(* IEC 61131-3 sources: DigitalTwin/sim-plc/plc, 2 files *)

(* ---- pump_station.st ---- *)
(*
  Pump station lead/lag control: OpenPLC Structured Text program.

  Specification: design/pump-station-design.md, section 4 (logic) and 5 (register map).

  Field I/O (%IX100, %QX100, %IW100) comes from the process simulator, which
  OpenPLC polls as a Modbus "slave device" (Generic TCP, 10.10.0.10:5020).
  The HMI reads the status block %QW0..%QW7 (holding registers 0..7) and
  writes settings to %MW0..%MW10 (holding registers 1024..1034).

  Pressures are UINT scaled x10: 1200 means 120.0 psi.

  Scan order, the same as every PLC: inputs are copied in, this program runs
  top to bottom once, outputs are copied out. Then it starts again.
*)
PROGRAM PumpStation
  VAR
    (* ---- Field inputs from the simulator (design 5.1) ---- *)
    P1_RUNNING    AT %IX100.0 : BOOL;
    P2_RUNNING    AT %IX100.1 : BOOL;
    P1_FAULT      AT %IX100.2 : BOOL;
    P2_FAULT      AT %IX100.3 : BOOL;
    PT101_DISCH   AT %IW100 : UINT;   (* discharge pressure, psi x10 *)
    PT100_SUCT    AT %IW101 : UINT;   (* suction pressure, psi x10 *)
    DEMAND        AT %IW102 : UINT;   (* pipeline demand, % x10 *)
    SIM_HEARTBEAT AT %IW103 : UINT;   (* +1 every simulator step *)

    (* ---- Field outputs to the simulator ---- *)
    P1_RUN_CMD AT %QX100.0 : BOOL;
    P2_RUN_CMD AT %QX100.1 : BOOL;

    (* ---- Status for the HMI: holding registers 0..7 (design 5.2) ---- *)
    HMI_DISCH_PRESS AT %QW0 : UINT;
    HMI_SUCT_PRESS  AT %QW1 : UINT;
    HMI_DEMAND      AT %QW2 : UINT;
    HMI_STATUS      AT %QW3 : UINT;
    HMI_ALARMS      AT %QW4 : UINT;
    HMI_LEAD_PUMP   AT %QW5 : UINT;
    HMI_MODE_ACTIVE AT %QW6 : UINT;
    PLC_HEARTBEAT   AT %QW7 : UINT;

    (* ---- Settings and commands from the HMI: holding registers 1024..1034 (design 5.3) ---- *)
    SP_PRESSURE     AT %MW0 : UINT;   (* lag start pressure, psi x10 *)
    SP_LAG_STOP     AT %MW1 : UINT;   (* lag stop pressure, psi x10 *)
    SP_LOW_ALARM    AT %MW2 : UINT;
    SP_HIGH_ALARM   AT %MW3 : UINT;
    LAG_START_DELAY AT %MW4 : UINT;   (* seconds *)
    LAG_STOP_DELAY  AT %MW5 : UINT;   (* seconds *)
    CMD_MODE        AT %MW6 : UINT;   (* 0 Off, 1 Auto, 2 Manual *)
    CMD_LEAD_SELECT AT %MW7 : UINT;   (* 1 = P1, 2 = P2 *)
    CMD_MANUAL_P1   AT %MW8 : UINT;   (* Manual mode: 1 run, 0 stop *)
    CMD_MANUAL_P2   AT %MW9 : UINT;
    CMD_ALARM_RESET AT %MW10 : UINT;  (* HMI writes 1; the PLC clears it *)
  END_VAR

  VAR
    (* Control state *)
    Mode       : UINT := 0;
    LastMode   : UINT := 0;
    ActiveLead : UINT := 1;        (* lead pump after any failover: 1 or 2 *)
    LagRun     : BOOL := FALSE;    (* Auto logic wants the lag pump running *)
    Handover   : BOOL := FALSE;    (* lead change in progress: keep the old lead on *)
    OldLead    : UINT := 0;
    P1Cmd      : BOOL := FALSE;
    P2Cmd      : BOOL := FALSE;
    LeadRunning : BOOL;
    LagAvail   : BOOL;
    LeadAvail  : BOOL;

    (* Pump failure latches: fault feedback or failed to start. A failed pump
       is locked out (never commanded) until the operator presses Reset and
       the simulator no longer reports a fault. *)
    P1Failed : BOOL := FALSE;
    P2Failed : BOOL := FALSE;
    P1StartTmr : TON;   (* run commanded but no running feedback *)
    P2StartTmr : TON;

    (* Lead/lag timers: the time delays that stop short-cycling *)
    LagStartTmr : TON;
    LagStopTmr  : TON;

    (* Alarms (design 4.3) *)
    LowArmTmr   : TON;   (* start-up bypass for the low-pressure alarm *)
    LowPressTmr : TON;
    HighPressTmr : TON;
    CommLossTmr : TON;
    LastSimHb   : UINT := 0;
    AlmLow   : BOOL := FALSE;
    AlmHigh  : BOOL := FALSE;
    AlmComm  : BOOL := FALSE;
    AlmUnack : BOOL := FALSE;
    AnyAlarm : BOOL;
    PrevAnyAlarm : BOOL := FALSE;
    ResetReq : BOOL;
    CommOk   : BOOL;
    LagRunning : BOOL;
  END_VAR

  (* =====================================================================
     1. First scan: load defaults (design 4.4).
        %MW memory is not kept across a runtime restart, so a zero setpoint
        means "never configured".
     ===================================================================== *)
  IF SP_PRESSURE = 0 THEN
    SP_PRESSURE     := 1200;   (* 120.0 psi *)
    SP_LAG_STOP     := 1450;   (* 145.0 psi *)
    SP_LOW_ALARM    := 1100;   (* 110.0 psi *)
    SP_HIGH_ALARM   := 1600;   (* 160.0 psi *)
    LAG_START_DELAY := 5;
    LAG_STOP_DELAY  := 30;
    CMD_MODE        := 1;      (* Auto *)
    CMD_LEAD_SELECT := 1;      (* P1 *)
    CMD_MANUAL_P1   := 0;
    CMD_MANUAL_P2   := 0;
    CMD_ALARM_RESET := 0;
  END_IF;

  (* =====================================================================
     2. Clamp HMI settings to their allowed ranges (design 5.3).
        The clamped value is written back, so the HMI reads back what the
        PLC is actually using.
     ===================================================================== *)
  SP_PRESSURE := LIMIT(800, SP_PRESSURE, 1500);
  IF SP_LAG_STOP < SP_PRESSURE + 100 THEN
    SP_LAG_STOP := SP_PRESSURE + 100;   (* hysteresis of at least 10 psi *)
  END_IF;
  LAG_START_DELAY := LIMIT(1, LAG_START_DELAY, 60);
  LAG_STOP_DELAY  := LIMIT(5, LAG_STOP_DELAY, 300);
  CMD_MODE        := MIN(CMD_MODE, 2);
  CMD_LEAD_SELECT := LIMIT(1, CMD_LEAD_SELECT, 2);
  CMD_MANUAL_P1   := MIN(CMD_MANUAL_P1, 1);
  CMD_MANUAL_P2   := MIN(CMD_MANUAL_P2, 1);
  Mode := CMD_MODE;

  ResetReq := CMD_ALARM_RESET <> 0;

  (* =====================================================================
     3. Pump health. Fault feedback, or no running feedback 5 s after a run
        command, fails the pump (design 4.2 step 4 and 4.3).
     ===================================================================== *)
  P1StartTmr(IN := P1_RUN_CMD AND NOT P1_RUNNING, PT := T#5s);
  P2StartTmr(IN := P2_RUN_CMD AND NOT P2_RUNNING, PT := T#5s);
  IF P1_FAULT OR P1StartTmr.Q THEN P1Failed := TRUE; END_IF;
  IF P2_FAULT OR P2StartTmr.Q THEN P2Failed := TRUE; END_IF;
  IF ResetReq AND NOT P1_FAULT THEN P1Failed := FALSE; END_IF;
  IF ResetReq AND NOT P2_FAULT THEN P2Failed := FALSE; END_IF;

  (* =====================================================================
     4. Pump control by mode (design 4.1, 4.2)
     ===================================================================== *)
  IF Mode = 1 THEN
    (* ---------------- Auto: lead/lag ---------------- *)

    (* Entering Auto: take the operator's lead choice, and keep whatever
       is already running so the switch causes no bump. *)
    IF LastMode <> 1 THEN
      ActiveLead := CMD_LEAD_SELECT;
      IF ActiveLead = 1 THEN LagRun := P2Cmd; ELSE LagRun := P1Cmd; END_IF;
      Handover := FALSE;
    END_IF;

    (* Failover: the lead pump has failed and the other one is healthy, so
       promote it. The HMI lead selection follows, so the station does not
       swap back on its own once the failed pump is reset. *)
    IF ((ActiveLead = 1) AND P1Failed AND NOT P2Failed) OR
       ((ActiveLead = 2) AND P2Failed AND NOT P1Failed) THEN
      ActiveLead := 3 - ActiveLead;
      CMD_LEAD_SELECT := ActiveLead;
      LagRun := FALSE;
      Handover := FALSE;
    END_IF;

    (* Operator changed the lead pump: applied only while the lag pump is
       stopped (design 4.2 step 5). The old lead keeps running until the new
       one reports running, so pressure does not dip during the swap. *)
    IF (CMD_LEAD_SELECT <> ActiveLead) AND NOT LagRun AND NOT Handover THEN
      IF ((CMD_LEAD_SELECT = 1) AND NOT P1Failed) OR
         ((CMD_LEAD_SELECT = 2) AND NOT P2Failed) THEN
        OldLead := ActiveLead;
        ActiveLead := CMD_LEAD_SELECT;
        Handover := TRUE;
      END_IF;
    END_IF;

    IF ActiveLead = 1 THEN
      LeadAvail := NOT P1Failed;  LagAvail := NOT P2Failed;  LeadRunning := P1_RUNNING;
    ELSE
      LeadAvail := NOT P2Failed;  LagAvail := NOT P1Failed;  LeadRunning := P2_RUNNING;
    END_IF;

    IF Handover AND (LeadRunning OR NOT LeadAvail) THEN
      Handover := FALSE;
    END_IF;

    (* Lag start: pressure below setpoint for the start delay (step 2) *)
    LagStartTmr(IN := (PT101_DISCH < SP_PRESSURE) AND NOT LagRun AND LagAvail AND NOT Handover,
                PT := T#1s * UINT_TO_DINT(LAG_START_DELAY));
    IF LagStartTmr.Q THEN
      LagRun := TRUE;
    END_IF;

    (* Lag stop: pressure above the lag stop pressure for the stop delay (step 3).
       The gap between 120 and 145 psi is the hysteresis that stops cycling. *)
    LagStopTmr(IN := LagRun AND (PT101_DISCH > SP_LAG_STOP),
               PT := T#1s * UINT_TO_DINT(LAG_STOP_DELAY));
    IF LagStopTmr.Q OR NOT LagAvail THEN
      LagRun := FALSE;
    END_IF;

    (* Lead always runs (step 1); lag runs when called for *)
    IF ActiveLead = 1 THEN
      P1Cmd := TRUE;
      P2Cmd := LagRun OR (Handover AND OldLead = 2);
    ELSE
      P2Cmd := TRUE;
      P1Cmd := LagRun OR (Handover AND OldLead = 1);
    END_IF;

  ELSIF Mode = 2 THEN
    (* ---------------- Manual: operator runs each pump ---------------- *)
    P1Cmd := CMD_MANUAL_P1 = 1;
    P2Cmd := CMD_MANUAL_P2 = 1;
    LagRun := FALSE;
    Handover := FALSE;

  ELSE
    (* ---------------- Off ---------------- *)
    P1Cmd := FALSE;
    P2Cmd := FALSE;
    LagRun := FALSE;
    Handover := FALSE;
  END_IF;

  (* Interlock in every mode: a failed pump is never commanded *)
  IF P1Failed THEN P1Cmd := FALSE; END_IF;
  IF P2Failed THEN P2Cmd := FALSE; END_IF;
  P1_RUN_CMD := P1Cmd;
  P2_RUN_CMD := P2Cmd;

  (* Outside Manual, the manual commands track the pumps, so switching to
     Manual leaves them as they are (bumpless transfer). *)
  IF Mode <> 2 THEN
    CMD_MANUAL_P1 := BOOL_TO_UINT(P1Cmd);
    CMD_MANUAL_P2 := BOOL_TO_UINT(P2Cmd);
  END_IF;
  LastMode := Mode;

  (* =====================================================================
     5. Alarms (design 4.3). Each one latches until the operator presses
        Reset AND its condition has cleared.
     ===================================================================== *)

  (* Low pressure is armed once the station has been out of Off for 15 s,
     so a normal start-up (pressure rising from 20 psi) does not alarm. *)
  LowArmTmr(IN := Mode <> 0, PT := T#15s);
  LowPressTmr(IN := LowArmTmr.Q AND (PT101_DISCH < SP_LOW_ALARM), PT := T#5s);
  HighPressTmr(IN := PT101_DISCH > SP_HIGH_ALARM, PT := T#5s);

  (* Simulator comm loss: heartbeat has not changed for 3 s *)
  CommLossTmr(IN := SIM_HEARTBEAT = LastSimHb, PT := T#3s);
  LastSimHb := SIM_HEARTBEAT;
  CommOk := NOT CommLossTmr.Q;

  IF LowPressTmr.Q  THEN AlmLow  := TRUE; END_IF;
  IF HighPressTmr.Q THEN AlmHigh := TRUE; END_IF;
  IF CommLossTmr.Q  THEN AlmComm := TRUE; END_IF;

  IF ResetReq THEN
    IF NOT LowPressTmr.Q  THEN AlmLow  := FALSE; END_IF;
    IF NOT HighPressTmr.Q THEN AlmHigh := FALSE; END_IF;
    IF NOT CommLossTmr.Q  THEN AlmComm := FALSE; END_IF;
    AlmUnack := FALSE;          (* Reset also acknowledges *)
    CMD_ALARM_RESET := 0;       (* handled *)
  END_IF;

  (* A newly raised alarm is unacknowledged until the next Reset *)
  AnyAlarm := AlmLow OR AlmHigh OR P1Failed OR P2Failed OR AlmComm;
  IF AnyAlarm AND NOT PrevAnyAlarm THEN AlmUnack := TRUE; END_IF;
  PrevAnyAlarm := AnyAlarm;

  (* =====================================================================
     6. Status block for the HMI (design 5.2)
     ===================================================================== *)
  IF ActiveLead = 1 THEN LagRunning := P2_RUNNING; ELSE LagRunning := P1_RUNNING; END_IF;

  HMI_DISCH_PRESS := PT101_DISCH;
  HMI_SUCT_PRESS  := PT100_SUCT;
  HMI_DEMAND      := DEMAND;
  HMI_STATUS := BOOL_TO_UINT(P1_RUN_CMD)
              + BOOL_TO_UINT(P1_RUNNING) * 2
              + BOOL_TO_UINT(P2_RUN_CMD) * 4
              + BOOL_TO_UINT(P2_RUNNING) * 8
              + BOOL_TO_UINT(LagRunning) * 16
              + BOOL_TO_UINT(CommOk)     * 32;
  HMI_ALARMS := BOOL_TO_UINT(AlmLow)
              + BOOL_TO_UINT(AlmHigh)  * 2
              + BOOL_TO_UINT(P1Failed) * 4
              + BOOL_TO_UINT(P2Failed) * 8
              + BOOL_TO_UINT(AlmComm)  * 16
              + BOOL_TO_UINT(AlmUnack) * 32768;
  HMI_LEAD_PUMP   := ActiveLead;
  HMI_MODE_ACTIVE := Mode;

  IF PLC_HEARTBEAT = 65535 THEN
    PLC_HEARTBEAT := 0;
  ELSE
    PLC_HEARTBEAT := PLC_HEARTBEAT + 1;
  END_IF;
END_PROGRAM

CONFIGURATION Config0
  RESOURCE Res0 ON PLC
    TASK MainTask(INTERVAL := T#100ms, PRIORITY := 0);
    PROGRAM Inst0 WITH MainTask : PumpStation;
  END_RESOURCE
END_CONFIGURATION

(* ---- pump_station_ld.st ---- *)
(*
  Generated from the ladder program in pump_station_ld/plc.xml by OpenPLC Editor's
  code generator. Do not edit this file: change the ladder in OpenPLC Editor instead.

  Upload this file to OpenPLC Runtime (Programs -> Upload program), or run
      python3 deploy_to_openplc.py --program pump_station_ld.st
  It behaves exactly like pump_station.st and uses the same register map.
*)
PROGRAM PumpStation
  VAR
    LoadDefaults : BOOL;
    MinLagStop : UINT;
    ModeAuto : BOOL;
    ModeManual : BOOL;
    SelP2 : BOOL;
    ManP1 : BOOL;
    ManP2 : BOOL;
    ResetReq : BOOL;
    PressBelowSP : BOOL;
    PressAboveLagStop : BOOL;
    PressBelowLowAlm : BOOL;
    PressAboveHighAlm : BOOL;
    P1StartTmr : TON;
    P2StartTmr : TON;
    P1StartFail : BOOL;
    P2StartFail : BOOL;
    P1Failed : BOOL;
    P2Failed : BOOL;
    EnterAuto : BOOL;
    LeadIsP2 : BOOL;
    LagPumpCmd : BOOL;
    FailToP2 : BOOL;
    FailToP1 : BOOL;
    LeadChange : BOOL;
    LagRun : BOOL;
    Handover : BOOL;
    LeadAvail : BOOL;
    LagAvail : BOOL;
    LeadRunning : BOOL;
    LagStartPT : TIME;
    LagStopPT : TIME;
    LagStartTmr : TON;
    LagStopTmr : TON;
    LagStartDone : BOOL;
    LagStopDone : BOOL;
    LowArmTmr : TON;
    LowPressTmr : TON;
    HighPressTmr : TON;
    CommLossTmr : TON;
    LowArmed : BOOL;
    LowPressOn : BOOL;
    HighPressOn : BOOL;
    SimHbFrozen : BOOL;
    LastSimHb : UINT;
    CommLost : BOOL;
    CommOk : BOOL;
    AlmLow : BOOL;
    AlmHigh : BOOL;
    AlmComm : BOOL;
    AlmUnack : BOOL;
    AnyAlarm : BOOL;
    LagRunning : BOOL;
    StatusWord : UINT;
    AlarmWord : UINT;
    HbWrap : BOOL;
  END_VAR
  VAR
    P1_RUNNING AT %IX100.0 : BOOL;
    P2_RUNNING AT %IX100.1 : BOOL;
    P1_FAULT AT %IX100.2 : BOOL;
    P2_FAULT AT %IX100.3 : BOOL;
    PT101_DISCH AT %IW100 : UINT;
    PT100_SUCT AT %IW101 : UINT;
    DEMAND AT %IW102 : UINT;
    SIM_HEARTBEAT AT %IW103 : UINT;
    P1_RUN_CMD AT %QX100.0 : BOOL;
    P2_RUN_CMD AT %QX100.1 : BOOL;
    HMI_DISCH_PRESS AT %QW0 : UINT;
    HMI_SUCT_PRESS AT %QW1 : UINT;
    HMI_DEMAND AT %QW2 : UINT;
    HMI_STATUS AT %QW3 : UINT;
    HMI_ALARMS AT %QW4 : UINT;
    HMI_LEAD_PUMP AT %QW5 : UINT;
    HMI_MODE_ACTIVE AT %QW6 : UINT;
    PLC_HEARTBEAT AT %QW7 : UINT;
    SP_PRESSURE AT %MW0 : UINT;
    SP_LAG_STOP AT %MW1 : UINT;
    SP_LOW_ALARM AT %MW2 : UINT;
    SP_HIGH_ALARM AT %MW3 : UINT;
    LAG_START_DELAY AT %MW4 : UINT;
    LAG_STOP_DELAY AT %MW5 : UINT;
    CMD_MODE AT %MW6 : UINT;
    CMD_LEAD_SELECT AT %MW7 : UINT;
    CMD_MANUAL_P1 AT %MW8 : UINT;
    CMD_MANUAL_P2 AT %MW9 : UINT;
    CMD_ALARM_RESET AT %MW10 : UINT;
  END_VAR
  VAR
    _TMP_EQ5_OUT : BOOL;
    _TMP_MOVE11_ENO : BOOL;
    _TMP_MOVE11_OUT : UINT;
    _TMP_MOVE14_ENO : BOOL;
    _TMP_MOVE14_OUT : UINT;
    _TMP_MOVE17_ENO : BOOL;
    _TMP_MOVE17_OUT : UINT;
    _TMP_MOVE20_ENO : BOOL;
    _TMP_MOVE20_OUT : UINT;
    _TMP_MOVE23_ENO : BOOL;
    _TMP_MOVE23_OUT : UINT;
    _TMP_MOVE26_ENO : BOOL;
    _TMP_MOVE26_OUT : UINT;
    _TMP_MOVE29_ENO : BOOL;
    _TMP_MOVE29_OUT : UINT;
    _TMP_MOVE32_ENO : BOOL;
    _TMP_MOVE32_OUT : UINT;
    _TMP_MOVE35_ENO : BOOL;
    _TMP_MOVE35_OUT : UINT;
    _TMP_MOVE38_ENO : BOOL;
    _TMP_MOVE38_OUT : UINT;
    _TMP_MOVE41_ENO : BOOL;
    _TMP_MOVE41_OUT : UINT;
    _TMP_LIMIT48_ENO : BOOL;
    _TMP_LIMIT48_OUT : UINT;
    _TMP_ADD53_ENO : BOOL;
    _TMP_ADD53_OUT : UINT;
    _TMP_MAX58_ENO : BOOL;
    _TMP_MAX58_OUT : UINT;
    _TMP_LIMIT64_ENO : BOOL;
    _TMP_LIMIT64_OUT : UINT;
    _TMP_LIMIT70_ENO : BOOL;
    _TMP_LIMIT70_OUT : UINT;
    _TMP_MIN76_ENO : BOOL;
    _TMP_MIN76_OUT : UINT;
    _TMP_LIMIT82_ENO : BOOL;
    _TMP_LIMIT82_OUT : UINT;
    _TMP_MIN87_ENO : BOOL;
    _TMP_MIN87_OUT : UINT;
    _TMP_MIN92_ENO : BOOL;
    _TMP_MIN92_OUT : UINT;
    _TMP_EQ98_OUT : BOOL;
    _TMP_EQ102_OUT : BOOL;
    _TMP_EQ107_OUT : BOOL;
    _TMP_EQ111_OUT : BOOL;
    _TMP_EQ115_OUT : BOOL;
    _TMP_NE119_OUT : BOOL;
    _TMP_LT124_OUT : BOOL;
    _TMP_GT128_OUT : BOOL;
    _TMP_LT132_OUT : BOOL;
    _TMP_GT136_OUT : BOOL;
    R_TRIG1 : R_TRIG;
    _TMP_MOVE220_ENO : BOOL;
    _TMP_MOVE220_OUT : UINT;
    _TMP_MOVE227_ENO : BOOL;
    _TMP_MOVE227_OUT : UINT;
    _TMP_UINT_TO_TIME286_ENO : BOOL;
    _TMP_UINT_TO_TIME286_OUT : TIME;
    _TMP_UINT_TO_TIME290_ENO : BOOL;
    _TMP_UINT_TO_TIME290_OUT : TIME;
    _TMP_BOOL_TO_UINT352_ENO : BOOL;
    _TMP_BOOL_TO_UINT352_OUT : UINT;
    _TMP_BOOL_TO_UINT355_ENO : BOOL;
    _TMP_BOOL_TO_UINT355_OUT : UINT;
    _TMP_EQ382_OUT : BOOL;
    _TMP_MOVE390_ENO : BOOL;
    _TMP_MOVE390_OUT : UINT;
    _TMP_MOVE417_ENO : BOOL;
    _TMP_MOVE417_OUT : UINT;
    R_TRIG2 : R_TRIG;
    _TMP_MOVE445_ENO : BOOL;
    _TMP_MOVE445_OUT : UINT;
    _TMP_MOVE449_ENO : BOOL;
    _TMP_MOVE449_OUT : UINT;
    _TMP_MOVE453_ENO : BOOL;
    _TMP_MOVE453_OUT : UINT;
    _TMP_SEL459_ENO : BOOL;
    _TMP_SEL459_OUT : UINT;
    _TMP_MOVE463_ENO : BOOL;
    _TMP_MOVE463_OUT : UINT;
    _TMP_MOVE468_ENO : BOOL;
    _TMP_MOVE468_OUT : UINT;
    _TMP_ADD475_ENO : BOOL;
    _TMP_ADD475_OUT : UINT;
    _TMP_ADD481_ENO : BOOL;
    _TMP_ADD481_OUT : UINT;
    _TMP_ADD487_ENO : BOOL;
    _TMP_ADD487_OUT : UINT;
    _TMP_ADD493_ENO : BOOL;
    _TMP_ADD493_OUT : UINT;
    _TMP_ADD499_ENO : BOOL;
    _TMP_ADD499_OUT : UINT;
    _TMP_ADD505_ENO : BOOL;
    _TMP_ADD505_OUT : UINT;
    _TMP_MOVE508_ENO : BOOL;
    _TMP_MOVE508_OUT : UINT;
    _TMP_MOVE513_ENO : BOOL;
    _TMP_MOVE513_OUT : UINT;
    _TMP_ADD520_ENO : BOOL;
    _TMP_ADD520_OUT : UINT;
    _TMP_ADD526_ENO : BOOL;
    _TMP_ADD526_OUT : UINT;
    _TMP_ADD532_ENO : BOOL;
    _TMP_ADD532_OUT : UINT;
    _TMP_ADD538_ENO : BOOL;
    _TMP_ADD538_OUT : UINT;
    _TMP_ADD544_ENO : BOOL;
    _TMP_ADD544_OUT : UINT;
    _TMP_ADD550_ENO : BOOL;
    _TMP_ADD550_OUT : UINT;
    _TMP_MOVE553_ENO : BOOL;
    _TMP_MOVE553_OUT : UINT;
    _TMP_EQ559_OUT : BOOL;
    _TMP_ADD565_ENO : BOOL;
    _TMP_ADD565_OUT : UINT;
    _TMP_MOVE570_ENO : BOOL;
    _TMP_MOVE570_OUT : UINT;
  END_VAR

  _TMP_EQ5_OUT := EQ(SP_PRESSURE, 0);
  LoadDefaults := _TMP_EQ5_OUT;
  _TMP_MOVE11_OUT := MOVE(EN := LoadDefaults, IN := 1200, ENO => _TMP_MOVE11_ENO);
  IF _TMP_MOVE11_ENO THEN
      SP_PRESSURE := _TMP_MOVE11_OUT;
  END_IF;
  _TMP_MOVE14_OUT := MOVE(EN := LoadDefaults, IN := 1450, ENO => _TMP_MOVE14_ENO);
  IF _TMP_MOVE14_ENO THEN
      SP_LAG_STOP := _TMP_MOVE14_OUT;
  END_IF;
  _TMP_MOVE17_OUT := MOVE(EN := LoadDefaults, IN := 1100, ENO => _TMP_MOVE17_ENO);
  IF _TMP_MOVE17_ENO THEN
      SP_LOW_ALARM := _TMP_MOVE17_OUT;
  END_IF;
  _TMP_MOVE20_OUT := MOVE(EN := LoadDefaults, IN := 1600, ENO => _TMP_MOVE20_ENO);
  IF _TMP_MOVE20_ENO THEN
      SP_HIGH_ALARM := _TMP_MOVE20_OUT;
  END_IF;
  _TMP_MOVE23_OUT := MOVE(EN := LoadDefaults, IN := 5, ENO => _TMP_MOVE23_ENO);
  IF _TMP_MOVE23_ENO THEN
      LAG_START_DELAY := _TMP_MOVE23_OUT;
  END_IF;
  _TMP_MOVE26_OUT := MOVE(EN := LoadDefaults, IN := 30, ENO => _TMP_MOVE26_ENO);
  IF _TMP_MOVE26_ENO THEN
      LAG_STOP_DELAY := _TMP_MOVE26_OUT;
  END_IF;
  _TMP_MOVE29_OUT := MOVE(EN := LoadDefaults, IN := 1, ENO => _TMP_MOVE29_ENO);
  IF _TMP_MOVE29_ENO THEN
      CMD_MODE := _TMP_MOVE29_OUT;
  END_IF;
  _TMP_MOVE32_OUT := MOVE(EN := LoadDefaults, IN := 1, ENO => _TMP_MOVE32_ENO);
  IF _TMP_MOVE32_ENO THEN
      CMD_LEAD_SELECT := _TMP_MOVE32_OUT;
  END_IF;
  _TMP_MOVE35_OUT := MOVE(EN := LoadDefaults, IN := 0, ENO => _TMP_MOVE35_ENO);
  IF _TMP_MOVE35_ENO THEN
      CMD_MANUAL_P1 := _TMP_MOVE35_OUT;
  END_IF;
  _TMP_MOVE38_OUT := MOVE(EN := LoadDefaults, IN := 0, ENO => _TMP_MOVE38_ENO);
  IF _TMP_MOVE38_ENO THEN
      CMD_MANUAL_P2 := _TMP_MOVE38_OUT;
  END_IF;
  _TMP_MOVE41_OUT := MOVE(EN := LoadDefaults, IN := 0, ENO => _TMP_MOVE41_ENO);
  IF _TMP_MOVE41_ENO THEN
      CMD_ALARM_RESET := _TMP_MOVE41_OUT;
  END_IF;
  _TMP_LIMIT48_OUT := LIMIT(EN := TRUE, MN := 800, IN := SP_PRESSURE, MX := 1500, ENO => _TMP_LIMIT48_ENO);
  IF _TMP_LIMIT48_ENO THEN
      SP_PRESSURE := _TMP_LIMIT48_OUT;
  END_IF;
  _TMP_ADD53_OUT := ADD(EN := TRUE, IN1 := SP_PRESSURE, IN2 := 100, ENO => _TMP_ADD53_ENO);
  IF _TMP_ADD53_ENO THEN
      MinLagStop := _TMP_ADD53_OUT;
  END_IF;
  _TMP_MAX58_OUT := MAX(EN := TRUE, IN1 := SP_LAG_STOP, IN2 := MinLagStop, ENO => _TMP_MAX58_ENO);
  IF _TMP_MAX58_ENO THEN
      SP_LAG_STOP := _TMP_MAX58_OUT;
  END_IF;
  _TMP_LIMIT64_OUT := LIMIT(EN := TRUE, MN := 1, IN := LAG_START_DELAY, MX := 60, ENO => _TMP_LIMIT64_ENO);
  IF _TMP_LIMIT64_ENO THEN
      LAG_START_DELAY := _TMP_LIMIT64_OUT;
  END_IF;
  _TMP_LIMIT70_OUT := LIMIT(EN := TRUE, MN := 5, IN := LAG_STOP_DELAY, MX := 300, ENO => _TMP_LIMIT70_ENO);
  IF _TMP_LIMIT70_ENO THEN
      LAG_STOP_DELAY := _TMP_LIMIT70_OUT;
  END_IF;
  _TMP_MIN76_OUT := MIN(EN := TRUE, IN1 := CMD_MODE, IN2 := 2, ENO => _TMP_MIN76_ENO);
  IF _TMP_MIN76_ENO THEN
      CMD_MODE := _TMP_MIN76_OUT;
  END_IF;
  _TMP_LIMIT82_OUT := LIMIT(EN := TRUE, MN := 1, IN := CMD_LEAD_SELECT, MX := 2, ENO => _TMP_LIMIT82_ENO);
  IF _TMP_LIMIT82_ENO THEN
      CMD_LEAD_SELECT := _TMP_LIMIT82_OUT;
  END_IF;
  _TMP_MIN87_OUT := MIN(EN := TRUE, IN1 := CMD_MANUAL_P1, IN2 := 1, ENO => _TMP_MIN87_ENO);
  IF _TMP_MIN87_ENO THEN
      CMD_MANUAL_P1 := _TMP_MIN87_OUT;
  END_IF;
  _TMP_MIN92_OUT := MIN(EN := TRUE, IN1 := CMD_MANUAL_P2, IN2 := 1, ENO => _TMP_MIN92_ENO);
  IF _TMP_MIN92_ENO THEN
      CMD_MANUAL_P2 := _TMP_MIN92_OUT;
  END_IF;
  _TMP_EQ98_OUT := EQ(CMD_MODE, 1);
  ModeAuto := _TMP_EQ98_OUT;
  _TMP_EQ102_OUT := EQ(CMD_MODE, 2);
  ModeManual := _TMP_EQ102_OUT;
  _TMP_EQ107_OUT := EQ(CMD_LEAD_SELECT, 2);
  SelP2 := _TMP_EQ107_OUT;
  _TMP_EQ111_OUT := EQ(CMD_MANUAL_P1, 1);
  ManP1 := _TMP_EQ111_OUT;
  _TMP_EQ115_OUT := EQ(CMD_MANUAL_P2, 1);
  ManP2 := _TMP_EQ115_OUT;
  _TMP_NE119_OUT := NE(CMD_ALARM_RESET, 0);
  ResetReq := _TMP_NE119_OUT;
  _TMP_LT124_OUT := LT(PT101_DISCH, SP_PRESSURE);
  PressBelowSP := _TMP_LT124_OUT;
  _TMP_GT128_OUT := GT(PT101_DISCH, SP_LAG_STOP);
  PressAboveLagStop := _TMP_GT128_OUT;
  _TMP_LT132_OUT := LT(PT101_DISCH, SP_LOW_ALARM);
  PressBelowLowAlm := _TMP_LT132_OUT;
  _TMP_GT136_OUT := GT(PT101_DISCH, SP_HIGH_ALARM);
  PressAboveHighAlm := _TMP_GT136_OUT;
  P1StartTmr(IN := NOT(P1_RUNNING) AND P1_RUN_CMD, PT := T#5s);
  P1StartFail := P1StartTmr.Q;
  P2StartTmr(IN := NOT(P2_RUNNING) AND P2_RUN_CMD, PT := T#5s);
  P2StartFail := P2StartTmr.Q;
  IF P1StartFail OR P1_FAULT THEN
    P1Failed := TRUE; (*set*)
  END_IF;
  IF P2StartFail OR P2_FAULT THEN
    P2Failed := TRUE; (*set*)
  END_IF;
  IF NOT(P1_FAULT) AND ResetReq THEN
    P1Failed := FALSE; (*reset*)
  END_IF;
  IF NOT(P2_FAULT) AND ResetReq THEN
    P2Failed := FALSE; (*reset*)
  END_IF;
  R_TRIG1(CLK := ModeAuto);
  EnterAuto := R_TRIG1.Q;
  IF SelP2 AND EnterAuto THEN
    LeadIsP2 := TRUE; (*set*)
  END_IF;
  IF NOT(SelP2) AND EnterAuto THEN
    LeadIsP2 := FALSE; (*reset*)
  END_IF;
  LagPumpCmd := P1_RUN_CMD AND LeadIsP2 OR P2_RUN_CMD AND NOT(LeadIsP2);
  IF LagPumpCmd AND EnterAuto THEN
    LagRun := TRUE; (*set*)
  END_IF;
  IF NOT(LagPumpCmd) AND EnterAuto THEN
    LagRun := FALSE; (*reset*)
  END_IF;
  IF EnterAuto THEN
    Handover := FALSE; (*reset*)
  END_IF;
  FailToP2 := NOT(P2Failed) AND P1Failed AND NOT(LeadIsP2) AND ModeAuto;
  FailToP1 := NOT(P1Failed) AND P2Failed AND LeadIsP2 AND ModeAuto;
  IF FailToP2 THEN
    LeadIsP2 := TRUE; (*set*)
  END_IF;
  IF FailToP2 THEN
    SelP2 := TRUE; (*set*)
  END_IF;
  _TMP_MOVE220_OUT := MOVE(EN := FailToP2, IN := 2, ENO => _TMP_MOVE220_ENO);
  IF _TMP_MOVE220_ENO THEN
      CMD_LEAD_SELECT := _TMP_MOVE220_OUT;
  END_IF;
  IF FailToP1 THEN
    LeadIsP2 := FALSE; (*reset*)
  END_IF;
  IF FailToP1 THEN
    SelP2 := FALSE; (*reset*)
  END_IF;
  _TMP_MOVE227_OUT := MOVE(EN := FailToP1, IN := 1, ENO => _TMP_MOVE227_ENO);
  IF _TMP_MOVE227_ENO THEN
      CMD_LEAD_SELECT := _TMP_MOVE227_OUT;
  END_IF;
  IF FailToP1 OR FailToP2 THEN
    LagRun := FALSE; (*reset*)
  END_IF;
  IF FailToP1 OR FailToP2 THEN
    Handover := FALSE; (*reset*)
  END_IF;
  LeadChange := (NOT(P2Failed) AND NOT(LeadIsP2) AND SelP2 OR NOT(P1Failed) AND LeadIsP2 AND NOT(SelP2)) AND NOT(Handover) AND NOT(LagRun) AND ModeAuto;
  IF SelP2 AND LeadChange THEN
    LeadIsP2 := TRUE; (*set*)
  END_IF;
  IF NOT(SelP2) AND LeadChange THEN
    LeadIsP2 := FALSE; (*reset*)
  END_IF;
  IF LeadChange THEN
    Handover := TRUE; (*set*)
  END_IF;
  LeadAvail := NOT(P1Failed) AND NOT(LeadIsP2) OR NOT(P2Failed) AND LeadIsP2;
  LagAvail := NOT(P2Failed) AND NOT(LeadIsP2) OR NOT(P1Failed) AND LeadIsP2;
  LeadRunning := P1_RUNNING AND NOT(LeadIsP2) OR P2_RUNNING AND LeadIsP2;
  IF (LeadRunning OR NOT(LeadAvail)) AND Handover AND ModeAuto THEN
    Handover := FALSE; (*reset*)
  END_IF;
  _TMP_UINT_TO_TIME286_OUT := UINT_TO_TIME(EN := TRUE, IN := LAG_START_DELAY, ENO => _TMP_UINT_TO_TIME286_ENO);
  IF _TMP_UINT_TO_TIME286_ENO THEN
      LagStartPT := _TMP_UINT_TO_TIME286_OUT;
  END_IF;
  _TMP_UINT_TO_TIME290_OUT := UINT_TO_TIME(EN := TRUE, IN := LAG_STOP_DELAY, ENO => _TMP_UINT_TO_TIME290_ENO);
  IF _TMP_UINT_TO_TIME290_ENO THEN
      LagStopPT := _TMP_UINT_TO_TIME290_OUT;
  END_IF;
  LagStartTmr(EN := ModeAuto, IN := NOT(Handover) AND LagAvail AND NOT(LagRun) AND PressBelowSP, PT := LagStartPT);
  LagStartDone := LagStartTmr.Q;
  IF LagStartDone AND ModeAuto THEN
    LagRun := TRUE; (*set*)
  END_IF;
  LagStopTmr(EN := ModeAuto, IN := PressAboveLagStop AND LagRun, PT := LagStopPT);
  LagStopDone := LagStopTmr.Q;
  IF (LagStopDone OR NOT(LagAvail)) AND ModeAuto THEN
    LagRun := FALSE; (*reset*)
  END_IF;
  IF NOT(ModeAuto) THEN
    LagRun := FALSE; (*reset*)
  END_IF;
  IF NOT(ModeAuto) THEN
    Handover := FALSE; (*reset*)
  END_IF;
  P1_RUN_CMD := ((Handover OR LagRun OR NOT(LeadIsP2)) AND ModeAuto OR ManP1 AND ModeManual) AND NOT(P1Failed);
  P2_RUN_CMD := ((Handover OR LagRun OR LeadIsP2) AND ModeAuto OR ManP2 AND ModeManual) AND NOT(P2Failed);
  _TMP_BOOL_TO_UINT352_OUT := BOOL_TO_UINT(EN := NOT(ModeManual), IN := P1_RUN_CMD, ENO => _TMP_BOOL_TO_UINT352_ENO);
  IF _TMP_BOOL_TO_UINT352_ENO THEN
      CMD_MANUAL_P1 := _TMP_BOOL_TO_UINT352_OUT;
  END_IF;
  _TMP_BOOL_TO_UINT355_OUT := BOOL_TO_UINT(EN := NOT(ModeManual), IN := P2_RUN_CMD, ENO => _TMP_BOOL_TO_UINT355_ENO);
  IF _TMP_BOOL_TO_UINT355_ENO THEN
      CMD_MANUAL_P2 := _TMP_BOOL_TO_UINT355_OUT;
  END_IF;
  LowArmTmr(IN := ModeAuto OR ModeManual, PT := T#15s);
  LowArmed := LowArmTmr.Q;
  LowPressTmr(IN := PressBelowLowAlm AND LowArmed, PT := T#5s);
  LowPressOn := LowPressTmr.Q;
  HighPressTmr(IN := PressAboveHighAlm, PT := T#5s);
  HighPressOn := HighPressTmr.Q;
  _TMP_EQ382_OUT := EQ(SIM_HEARTBEAT, LastSimHb);
  SimHbFrozen := _TMP_EQ382_OUT;
  CommLossTmr(IN := SimHbFrozen, PT := T#3s);
  CommLost := CommLossTmr.Q;
  _TMP_MOVE390_OUT := MOVE(EN := TRUE, IN := SIM_HEARTBEAT, ENO => _TMP_MOVE390_ENO);
  IF _TMP_MOVE390_ENO THEN
      LastSimHb := _TMP_MOVE390_OUT;
  END_IF;
  CommOk := NOT(CommLost);
  IF LowPressOn THEN
    AlmLow := TRUE; (*set*)
  END_IF;
  IF HighPressOn THEN
    AlmHigh := TRUE; (*set*)
  END_IF;
  IF CommLost THEN
    AlmComm := TRUE; (*set*)
  END_IF;
  IF NOT(LowPressOn) AND ResetReq THEN
    AlmLow := FALSE; (*reset*)
  END_IF;
  IF NOT(HighPressOn) AND ResetReq THEN
    AlmHigh := FALSE; (*reset*)
  END_IF;
  IF NOT(CommLost) AND ResetReq THEN
    AlmComm := FALSE; (*reset*)
  END_IF;
  IF ResetReq THEN
    AlmUnack := FALSE; (*reset*)
  END_IF;
  _TMP_MOVE417_OUT := MOVE(EN := ResetReq, IN := 0, ENO => _TMP_MOVE417_ENO);
  IF _TMP_MOVE417_ENO THEN
      CMD_ALARM_RESET := _TMP_MOVE417_OUT;
  END_IF;
  AnyAlarm := AlmComm OR AlmHigh OR AlmLow OR P1Failed OR P2Failed;
  R_TRIG2(CLK := AnyAlarm);
  IF R_TRIG2.Q THEN
    AlmUnack := TRUE; (*set*)
  END_IF;
  LagRunning := P1_RUNNING AND LeadIsP2 OR P2_RUNNING AND NOT(LeadIsP2);
  _TMP_MOVE445_OUT := MOVE(EN := TRUE, IN := PT101_DISCH, ENO => _TMP_MOVE445_ENO);
  IF _TMP_MOVE445_ENO THEN
      HMI_DISCH_PRESS := _TMP_MOVE445_OUT;
  END_IF;
  _TMP_MOVE449_OUT := MOVE(EN := TRUE, IN := PT100_SUCT, ENO => _TMP_MOVE449_ENO);
  IF _TMP_MOVE449_ENO THEN
      HMI_SUCT_PRESS := _TMP_MOVE449_OUT;
  END_IF;
  _TMP_MOVE453_OUT := MOVE(EN := TRUE, IN := DEMAND, ENO => _TMP_MOVE453_ENO);
  IF _TMP_MOVE453_ENO THEN
      HMI_DEMAND := _TMP_MOVE453_OUT;
  END_IF;
  _TMP_SEL459_OUT := SEL(EN := TRUE, G := LeadIsP2, IN0 := 1, IN1 := 2, ENO => _TMP_SEL459_ENO);
  IF _TMP_SEL459_ENO THEN
      HMI_LEAD_PUMP := _TMP_SEL459_OUT;
  END_IF;
  _TMP_MOVE463_OUT := MOVE(EN := TRUE, IN := CMD_MODE, ENO => _TMP_MOVE463_ENO);
  IF _TMP_MOVE463_ENO THEN
      HMI_MODE_ACTIVE := _TMP_MOVE463_OUT;
  END_IF;
  _TMP_MOVE468_OUT := MOVE(EN := TRUE, IN := 0, ENO => _TMP_MOVE468_ENO);
  IF _TMP_MOVE468_ENO THEN
      StatusWord := _TMP_MOVE468_OUT;
  END_IF;
  _TMP_ADD475_OUT := ADD(EN := P1_RUN_CMD, IN1 := StatusWord, IN2 := 1, ENO => _TMP_ADD475_ENO);
  IF _TMP_ADD475_ENO THEN
      StatusWord := _TMP_ADD475_OUT;
  END_IF;
  _TMP_ADD481_OUT := ADD(EN := P1_RUNNING, IN1 := StatusWord, IN2 := 2, ENO => _TMP_ADD481_ENO);
  IF _TMP_ADD481_ENO THEN
      StatusWord := _TMP_ADD481_OUT;
  END_IF;
  _TMP_ADD487_OUT := ADD(EN := P2_RUN_CMD, IN1 := StatusWord, IN2 := 4, ENO => _TMP_ADD487_ENO);
  IF _TMP_ADD487_ENO THEN
      StatusWord := _TMP_ADD487_OUT;
  END_IF;
  _TMP_ADD493_OUT := ADD(EN := P2_RUNNING, IN1 := StatusWord, IN2 := 8, ENO => _TMP_ADD493_ENO);
  IF _TMP_ADD493_ENO THEN
      StatusWord := _TMP_ADD493_OUT;
  END_IF;
  _TMP_ADD499_OUT := ADD(EN := LagRunning, IN1 := StatusWord, IN2 := 16, ENO => _TMP_ADD499_ENO);
  IF _TMP_ADD499_ENO THEN
      StatusWord := _TMP_ADD499_OUT;
  END_IF;
  _TMP_ADD505_OUT := ADD(EN := CommOk, IN1 := StatusWord, IN2 := 32, ENO => _TMP_ADD505_ENO);
  IF _TMP_ADD505_ENO THEN
      StatusWord := _TMP_ADD505_OUT;
  END_IF;
  _TMP_MOVE508_OUT := MOVE(EN := TRUE, IN := StatusWord, ENO => _TMP_MOVE508_ENO);
  IF _TMP_MOVE508_ENO THEN
      HMI_STATUS := _TMP_MOVE508_OUT;
  END_IF;
  _TMP_MOVE513_OUT := MOVE(EN := TRUE, IN := 0, ENO => _TMP_MOVE513_ENO);
  IF _TMP_MOVE513_ENO THEN
      AlarmWord := _TMP_MOVE513_OUT;
  END_IF;
  _TMP_ADD520_OUT := ADD(EN := AlmLow, IN1 := AlarmWord, IN2 := 1, ENO => _TMP_ADD520_ENO);
  IF _TMP_ADD520_ENO THEN
      AlarmWord := _TMP_ADD520_OUT;
  END_IF;
  _TMP_ADD526_OUT := ADD(EN := AlmHigh, IN1 := AlarmWord, IN2 := 2, ENO => _TMP_ADD526_ENO);
  IF _TMP_ADD526_ENO THEN
      AlarmWord := _TMP_ADD526_OUT;
  END_IF;
  _TMP_ADD532_OUT := ADD(EN := P1Failed, IN1 := AlarmWord, IN2 := 4, ENO => _TMP_ADD532_ENO);
  IF _TMP_ADD532_ENO THEN
      AlarmWord := _TMP_ADD532_OUT;
  END_IF;
  _TMP_ADD538_OUT := ADD(EN := P2Failed, IN1 := AlarmWord, IN2 := 8, ENO => _TMP_ADD538_ENO);
  IF _TMP_ADD538_ENO THEN
      AlarmWord := _TMP_ADD538_OUT;
  END_IF;
  _TMP_ADD544_OUT := ADD(EN := AlmComm, IN1 := AlarmWord, IN2 := 16, ENO => _TMP_ADD544_ENO);
  IF _TMP_ADD544_ENO THEN
      AlarmWord := _TMP_ADD544_OUT;
  END_IF;
  _TMP_ADD550_OUT := ADD(EN := AlmUnack, IN1 := AlarmWord, IN2 := 32768, ENO => _TMP_ADD550_ENO);
  IF _TMP_ADD550_ENO THEN
      AlarmWord := _TMP_ADD550_OUT;
  END_IF;
  _TMP_MOVE553_OUT := MOVE(EN := TRUE, IN := AlarmWord, ENO => _TMP_MOVE553_ENO);
  IF _TMP_MOVE553_ENO THEN
      HMI_ALARMS := _TMP_MOVE553_OUT;
  END_IF;
  _TMP_EQ559_OUT := EQ(PLC_HEARTBEAT, 65535);
  HbWrap := _TMP_EQ559_OUT;
  _TMP_ADD565_OUT := ADD(EN := NOT(HbWrap), IN1 := PLC_HEARTBEAT, IN2 := 1, ENO => _TMP_ADD565_ENO);
  IF _TMP_ADD565_ENO THEN
      PLC_HEARTBEAT := _TMP_ADD565_OUT;
  END_IF;
  _TMP_MOVE570_OUT := MOVE(EN := HbWrap, IN := 0, ENO => _TMP_MOVE570_ENO);
  IF _TMP_MOVE570_ENO THEN
      PLC_HEARTBEAT := _TMP_MOVE570_OUT;
  END_IF;
END_PROGRAM

CONFIGURATION Config0

  RESOURCE Res0 ON PLC
    TASK MainTask(INTERVAL := T#100ms,PRIORITY := 0);
    PROGRAM Inst0 WITH MainTask : PumpStation;
  END_RESOURCE
END_CONFIGURATION
